FUNCTION F_OpcUaCreateObjectId (* Creates an OPC UA identifier for an object node type *)
  (* Standard: 61499-2; Description: Copyright (c) 2026 Monika Wenger This program and the accompanying materials are made available under the terms of the Eclipse Public License 2.0 which is available at https://www.eclipse.org/legal/epl-2.0/ SPDX-License-Identifier: EPL-2.0 *)
  (* Version 3.0, 2026-10-14, Monika Wenger *)
  PACKAGE eclipse4diac::opcua;
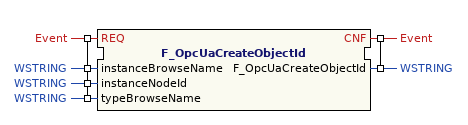
  EVENT_INPUT
    REQ WITH instanceBrowseName, instanceNodeId, typeBrowseName;
  END_EVENT
  EVENT_OUTPUT
    CNF WITH F_OpcUaCreateObjectId;
  END_EVENT
  VAR_INPUT
    instanceBrowseName : WSTRING;
    instanceNodeId : WSTRING;
    typeBrowseName : WSTRING;
  END_VAR
  VAR_OUTPUT
    F_OpcUaCreateObjectId : WSTRING;
  END_VAR
  BODY IN ST:
PACKAGE eclipse4diac::opcua;

(* Creates an OPC UA identifier for an object node type *)
FUNCTION F_OpcUaCreateObjectId : WSTRING
VAR_INPUT
	instanceBrowseName : WSTRING;
	instanceNodeId : WSTRING;
	typeBrowseName : WSTRING;
END_VAR
VAR CONSTANT
	PREFIX : WSTRING := "opc_ua[CREATE_OBJECT;";
	NODEID_TYPE : WSTRING := ",s=";
	SUFFIX : WSTRING := "]";
	SEPARATOR_PAIR : WSTRING := ";";
END_VAR
F_OpcUaCreateObjectId := CONCAT(PREFIX, typeBrowseName, SEPARATOR_PAIR, instanceBrowseName, NODEID_TYPE, instanceNodeId,
	SUFFIX);
END_FUNCTION
  END_BODY
END_FUNCTION
